ADAPTER buttons_automatic (* Adapter Interface *)
  (* Standard: 61499-1 *)
  (* Version 0.0, 10/22/2026, macie, Schneider Electric *)
  PACKAGE Main;
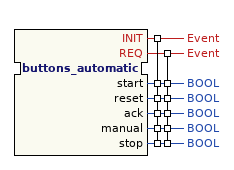
  EVENT_OUTPUT
    INIT WITH start, reset, ack, manual, stop;
    REQ WITH start, reset, ack, manual, stop;
  END_EVENT
  VAR_OUTPUT
    start : BOOL;
    reset : BOOL;
    ack : BOOL;
    manual : BOOL;
    stop : BOOL;
  END_VAR
  SERVICE SOCKET/PLUG
    SEQUENCE request_confirm
      SOCKET.REQ(start) -> PLUG.REQ(start);
      PLUG.CNF(CNFD) -> SOCKET.CNF(CNFD);
    END_SEQUENCE
    SEQUENCE indication_response
      PLUG.IND(INDD) -> SOCKET.IND(INDD);
      SOCKET.RSP(reset) -> PLUG.RSP(reset);
    END_SEQUENCE
  END_SERVICE
END_ADAPTER
